{region 'Documentation'}
(*!
<summary>Checks stable insertion into two slots, including a temporary gap before Finalize.</summary>
<description>Child mocks are inert interface identities and slot storage only; no child initialization or FB call is performed.</description>
*)
{endregion}
FUNCTION_BLOCK Test_RunControlBuilderSlotInsertion EXTENDS TestCaseBase
VAR
    FBuilder : RunControlConfigurationBuilder;
    FSuites : ARRAY[1..4] OF I_TestSuite;
    FChildA : TestSuiteMock;
    FChildB : TestSuiteMock;
    FChildC : TestSuiteMock;
    FChildD : TestSuiteMock;
    FScenarioExecuted : BOOL;
    FChecksEvaluated : BOOL;
    FRegistration : AssertTrue;
    FRegistrationMatches : BOOL;
    FOrder : AssertTrue;
    FOrderMatches : BOOL;
    FSlots : AssertTrue;
    FSlotsMatches : BOOL;
    FFinalization : AssertTrue;
    FFinalizationMatches : BOOL;
END_VAR

SUPER^();

{region 'Documentation'}
(*!
<summary>Contributes each owned Assertion once without executing it.</summary>
*)
{endregion}
METHOD PROTECTED AggregateResults
VAR_INPUT
    Aggregator : I_ResultAggregator; //! Borrowed result sink owned by the outer Test Case; add this test's checking Assertions without resetting or retaining the sink.
END_VAR
Aggregator.AddProvider(Provider := FRegistration);
Aggregator.AddProvider(Provider := FOrder);
Aggregator.AddProvider(Provider := FSlots);
Aggregator.AddProvider(Provider := FFinalization);
END_METHOD

{region 'Documentation'}
(*!
<summary>Requires successful base and owned Assertion initialization.</summary>
*)
{endregion}
METHOD PROTECTED CheckInitialization : BOOL //! TRUE when the inherited initialization check and this concrete fixture check both accept the setup.
CheckInitialization := FALSE;
IF NOT SUPER^.CheckInitialization() THEN
    RETURN;
END_IF;

CheckInitialization := FRegistration.IsInitialized
    AND FOrder.IsInitialized
    AND FSlots.IsInitialized
    AND FFinalization.IsInitialized;
END_METHOD

{region 'Documentation'}
(*!
<summary>Configures one direct builder scenario and its named Assertions.</summary>
*)
{endregion}
METHOD PROTECTED Configure
FPreparationStateCount := 0;
FTestStateCount := 1;
FScenarioExecuted := FALSE;
FChecksEvaluated := FALSE;

FRegistrationMatches := FALSE;
FRegistration.Initialize(Parent := THIS^,
    AssertionName := 'Registration');
FOrderMatches := FALSE;
FOrder.Initialize(Parent := THIS^,
    AssertionName := 'Order');
FSlotsMatches := FALSE;
FSlots.Initialize(Parent := THIS^,
    AssertionName := 'Slots');
FFinalizationMatches := FALSE;
FFinalization.Initialize(Parent := THIS^,
    AssertionName := 'Finalization');
END_METHOD

{region 'Documentation'}
(*!
<summary>Completes Abort immediately; no asynchronous resource operation is started.</summary>
*)
{endregion}
METHOD PROTECTED ProcessAbort
VAR_INPUT
    Enable : BOOL; //! Phase permission supplied by the owning Test Case; FALSE does not authorize progression, while observation may continue.
END_VAR
IF Enable THEN
    CompleteAbort();
END_IF;
END_METHOD

{region 'Documentation'}
(*!
<summary>Evaluates recorded observations and consumes pending resets on disabled calls.</summary>
*)
{endregion}
METHOD PROTECTED ProcessAssertions
VAR_INPUT
    Enable : BOOL; //! Phase permission supplied by the owning Test Case; FALSE does not authorize progression, while observation may continue.
END_VAR
FRegistration(Enable := Enable,
    State := State,
    IN := FRegistrationMatches);

FOrder(Enable := Enable,
    State := State,
    IN := FOrderMatches);

FSlots(Enable := Enable,
    State := State,
    IN := FSlotsMatches);

FFinalization(Enable := Enable,
    State := State,
    IN := FFinalizationMatches);

IF Enable AND FRegistration.EvaluationActive
    AND FOrder.EvaluationActive
    AND FSlots.EvaluationActive
    AND FFinalization.EvaluationActive THEN
    FChecksEvaluated := TRUE;
END_IF;
END_METHOD

{region 'Documentation'}
(*!
<summary>No Preparation phase is needed for synchronous builder calls.</summary>
*)
{endregion}
METHOD PROTECTED ProcessPreparations
VAR_INPUT
    // SA0033: Required override signature; this scenario has no Preparation work.
    {attribute 'analysis' := '-33'}
    Enable : BOOL; //! Phase permission supplied by the owning Test Case; FALSE does not authorize progression, while observation may continue.
END_VAR
END_METHOD

{region 'Documentation'}
(*!
<summary>Clears recorded checks and Assertion results; each scenario initializes its own builder.</summary>
*)
{endregion}
METHOD PROTECTED ProcessReset
FScenarioExecuted := FALSE;
FChecksEvaluated := FALSE;
FRegistrationMatches := FALSE;
FRegistration.Reset();
FOrderMatches := FALSE;
FOrder.Reset();
FSlotsMatches := FALSE;
FSlots.Reset();
FFinalizationMatches := FALSE;
FFinalization.Reset();
CompleteReset();
END_METHOD

{region 'Documentation'}
(*!
<summary>Runs setup operations once, then completes after their observations have been evaluated.</summary>
*)
{endregion}
METHOD PROTECTED ProcessTests
VAR_INPUT
    Enable : BOOL; //! Phase permission supplied by the owning Test Case; FALSE does not authorize progression, while observation may continue.
END_VAR
IF NOT Enable THEN
    RETURN;
END_IF;

IF FChecksEvaluated THEN
    CompleteTests();
ELSIF NOT FScenarioExecuted THEN
    RunScenario();
    FScenarioExecuted := TRUE;
END_IF;
END_METHOD

{region 'Documentation'}
(*!
<summary>Checks stable insertion into two slots, including a temporary gap before Finalize.</summary>
*)
{endregion}
METHOD PRIVATE RunScenario
VAR
    ChildA : I_TestSuite;
    ChildB : I_TestSuite;
    ChildC : I_TestSuite;
    ChildD : I_TestSuite;
    AcceptedA : BOOL;
    AcceptedB : BOOL;
    AcceptedC : BOOL;
    AcceptedD : BOOL;
    Config : ST_TestSuiteCollectionConfig;
END_VAR
ChildA := FChildA;
ChildB := FChildB;
ChildC := FChildC;
ChildD := FChildD;
FBuilder.Initialize(Mode := E_OrchestrationMode.ParallelSlots,
    TestSuites := FSuites);
AcceptedA := FBuilder.RegisterWithSlot(TestSuite := ChildA,
    ExecutionSlot := 2);
AcceptedB := FBuilder.RegisterWithSlot(TestSuite := ChildB,
    ExecutionSlot := 1);
AcceptedC := FBuilder.RegisterWithSlot(TestSuite := ChildC,
    ExecutionSlot := 2);
AcceptedD := FBuilder.RegisterWithSlot(TestSuite := ChildD,
    ExecutionSlot := 1);
FRegistrationMatches := AcceptedA AND AcceptedB AND AcceptedC AND AcceptedD;
FOrderMatches := (FSuites[1] = ChildB) AND (FSuites[2] = ChildD)
    AND (FSuites[3] = ChildA) AND (FSuites[4] = ChildC);
FSlotsMatches := (FChildA.ExecutionSlot = 2) AND (FChildB.ExecutionSlot = 1)
    AND (FChildC.ExecutionSlot = 2) AND (FChildD.ExecutionSlot = 1);

Config := FBuilder.Finalize();
FFinalizationMatches := Config.IsValid AND FBuilder.IsValid AND FBuilder.IsFinalized
    AND (Config.FirstIndex = 1) AND (Config.LastIndex = 4) AND (Config.Count = 4)
    AND (Config.Mode = E_OrchestrationMode.ParallelSlots);
END_METHOD

END_FUNCTION_BLOCK

(* stored: Version 1.1.0.1
   POU Test_RunControlBuilderSlotInsertion: Id {e38f5bb9-77c6-4f51-ad04-797f6f41d43f}, SpecialFunc None
   Folder Internal: Id {00570001-0057-4057-8057-000000000021}
   Method AggregateResults: Id {00570001-0057-4057-8057-00000000001f}
   Method CheckInitialization: Id {00570001-0057-4057-8057-000000000018}
   Method Configure: Id {00570001-0057-4057-8057-000000000017}
   Method ProcessAbort: Id {00570001-0057-4057-8057-00000000001a}
   Method ProcessAssertions: Id {00570001-0057-4057-8057-00000000001e}
   Method ProcessPreparations: Id {00570001-0057-4057-8057-000000000019}
   Method ProcessReset: Id {00570001-0057-4057-8057-00000000001b}
   Method ProcessTests: Id {00570001-0057-4057-8057-00000000001c}
   Method RunScenario: Id {00570001-0057-4057-8057-00000000001d} *)
